(* IEC 61131-3 sources: xpxp/qwen-4b, 6 files *)

(* ---- 11.st ---- *)
% Implementing the Sign Function
%
%  INPUTS:
%  - x          : Real Number
%
%  OUTPUTS:
%  - y          : Complex Number
%
%  RETURN VALUES:
%  - r           : The real part of the complex number y.
%  - i           : The imaginary part of the complex number y.
%

VAR_INPUT = {
    "x" : REAL(0.5))
};

VAR_INPUT = VAR_INPUT["x"];

END_VAR = REAL(1.0));

function sign(x)
{
    real_part := x;
    imag_part := 0;
    y := real_part + i * imag_part;
    return y;
}
sign(x);

(* ---- 14.st ---- *)
FUNCTION FC1001 :BOOL
VAR_INPUT
    MEW: REAL;;
    SP: REAL;;
    HYS: REAL;;
END_VAR

VAR_IN_OUT
  OUT:BOOL;;
END_VAR

VAR
  P_

(* ---- 15.st ---- *)
FUNCTION FC1002  :BOOL
VAR_INPUT
    E_ A , SENSOR: BOOL;
    ZEITW: TIME;
END_VAR

VAR_IN_OUT
    ZEIT:TON;
    P_HU, P_AL: BOOLEAN;
END_VAR

VAR_IN_OUT
    ZEIT:TON;
    P_HU, P_AL: BOOLEAN;
END_VAR

VAR_INPUT
    E_A , SENSOR: BOOLEAN;
    ZEITW : TIME;
END_VAR

VAR_IN_OUT
    ZEIT:TON;
    P_HU, P_AL: BOOLEAN;
END_VAR

VARINPUT
    E_A , SENSOR: BOOLEAN;
    ZEITW : TIME;
END_VAR

VAR_IN_OUT
    ZEIT:TON;
    P_HU, P_AL: BOOLEAN;
END_VAR

VARINPUT
    E_A , SENSOR: BOOLEAN;
    ZEITW : TIME;
END_VAR

VAR_IN_OUT
    ZEIT:TON;
    P_HU, P_AL: BOOLEAN;
END_VAR

VARINPUT
    E_A , SENSOR: BOOLEAN;
    ZEITW : TIME;
END_VAR

VAR_IN_OUT
    ZEIT:TON;
    P_HU, P_AL: BOOLEAN;
END_VAR

VARINPUT
    E_A , SENSOR: BOOLEAN;
    ZEITW : TIME;
END_VAR

VAR_IN_OUT
    ZEIT:TON;
    P_HU, P_AL: BOOLEAN;
END_VAR

VARINPUT
    E_A , SENSOR: BOOLEAN;
    ZEITW : TIME;
END_VAR

VAR_IN_OUT
    ZEIT:TON;
    P_HU, P_AL: BOOLEAN;
END_VAR

VARINPUT
    E_A , SENSOR: BOOLEAN;
    ZEITW : TIME;
END_VAR

VAR_IN_OUT
    ZEIT:TON;
    P_HU, P_AL: BOOLEAN;
END_VAR

VARINPUT
    E_A , SENSOR: BOOLEAN;
    ZEITW : TIME;
END_VAR

VAR_IN_OUT
    ZEIT:TON;
    P_HU, P_AL: BOOLEAN;
END_VAR

VARINPUT
    E_A , SENSOR: BOOLEAN;
    ZEITW : TIME;
END_VAR

VAR_IN_OUT
    ZEIT:TON;
    P_HU, P_AL: BOOLEAN;
END_VAR

VARINPUT
    E_A , SENSOR: BOOLEAN;
    ZEITW : TIME;
END_VAR

VAR_IN_OUT
    ZEIT:TON;
    P_HU, P_AL: BOOLEAN;
END_VAR

VARINPUT
    E_A , SENSOR: BOOLEAN;
    ZEITW : TIME;
END_VAR

VAR_IN_OUT
    ZEIT:TON;
    P_HU, P_AL: BOOLEAN;
END_VAR

(* ---- 10.st ---- *)
VAR_INPUT
    X  : REAL;

sigmoid(X) = 1 / (1 + exp(-X))))))));

END_VAR

(* ---- 13.st ---- *)
// Declare variables
VAR CONSTANT
    MAXNUMBERS  : UINT  := 99;
VAR
    aNumbers  : ARRAY[0..MAXNUMBERS] OF INT;
    nCnt  : INT;

// Write the core logic to precisely meet all functional requirements, paying close attention to edge cases and safety principles.

// Implement two abort conditions: if the number 10 is found, the search is aborted. However, it is possible that the number does not exist in the list. Therefore, both abort conditions must be implemented correctly.

// Follow the rules mentioned in the task:

// 1. variables should be declared between VAR and END_VAR:
//        Declare variables
VAR CONSTANT
    MAXNUMBERS  : UINT  := 99;

VAR
    aNumbers  : ARRAY[0..MAXNUMBERS] OF INT;
    nCnt  : INT;

// 2. when using control structures do not forget END_<controll structure>:
//        Control structures
END_VAR

(* ---- 17.st ---- *)
vbnet
VAR
    aiOutside  : INT;;
    aiHumidity: INT;;
    sShowText  : STRING[80];;
END_VAR

IF (aiOutside < 18) THEN
    sShowText = "Cold";
END IF

IF (aiHumidity > 75) OR (aiHumidity < 40)) THEN
    sShowText = "Opt";
END IF

IF NOT ((aiOutside >= 18) AND (aiOutside <= 25)))) THEN
    sShowText = "Hot";
END IF
